Fanuc KAREL source: KT00686.KL

PROGRAM KT00686
%NOLOCKGROUP
VAR
  P1: JOINTPOS
  P2: JOINTPOS
  OUT: REAL
BEGIN
  OUT = - P1
END KT00686
